// TIA Portal V21 export
// export: Created 2026-10-23T20:42:44.5110947Z, ExportSetting WithDefaults, DisplayName Totally Integrated Automation Portal, DisplayVersion V21 Update 1, DisplayName SINAMICS Startdrive Advanced, DisplayVersion V21 HF2, DisplayName SINAMICS Startdrive G110M, G120, G120C, G120D, G120P, G115D, DisplayVersion V21 HF2, DisplayName SINAMICS Startdrive G130, G150, S120, S150, G200, G220, S200, S210, S220, Innomotics MVD, DisplayVersion V21 HF2, DisplayName STEP 7 Professional, DisplayVersion V21 Update 1, DisplayName STEP 7 Safety, DisplayVersion V21, DisplayName Tech WebApplication, DisplayVersion V21, DisplayName WinCC Basic/Comfort/Advanced, DisplayVersion V21 Update 1, DisplayName WinCC Unified, DisplayVersion V21 Update 1
FUNCTION_BLOCK "FB_LadOpenBranch"   // FB8, LAD
TITLE = LAD open branch and parallel coils
{ S7_Optimized_Access := 'TRUE' }
VERSION : 0.1
// stored: AutoNumber true, IsIECCheckEnabled false, IsRetainMemResEnabled false, MemoryReserve 100, SetENOAutomatically false, UDAEnableTagReadback false
   VAR_INPUT
      Start : Bool;   // Start command
      Stop : Bool;   // Stop command
   END_VAR
   VAR_OUTPUT
      CoilA : Bool;   // First parallel coil
      CoilB : Bool;   // Second parallel coil
      CoilC : Bool;   // Third parallel coil, only without stop
      BranchOut : Bool;   // Coil of the network with the open branch
      StopLatched : Bool;   // Set by the open branch when stop is pressed during start
   END_VAR
   VAR
      StartCount : Int;   // Number of cycles with start pressed
   END_VAR
BEGIN

REGION Network 1: Several coils in parallel
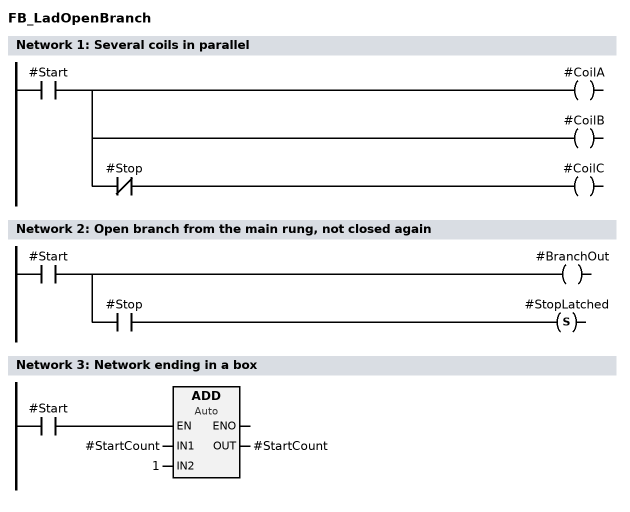
   RUNG wire#powerrail
      Contact( #Start )
      wire#w1
      Coil( #CoilA )
   END_RUNG
   RUNG wire#w1
      Coil( #CoilB )
   END_RUNG
   RUNG wire#w1
      I_Contact( #Stop )
      Coil( #CoilC )
   END_RUNG
   // the same network as SCL:
   #CoilA := #Start;
   #CoilB := #Start;
   #CoilC := #Start AND NOT #Stop;
END_REGION

REGION Network 2: Open branch from the main rung, not closed again
   RUNG wire#powerrail
      Contact( #Start )
      wire#w1
      Coil( #BranchOut )
   END_RUNG
   RUNG wire#w1
      Contact( #Stop )
      S_Coil( #StopLatched )
   END_RUNG
   // the same network as SCL:
   #BranchOut := #Start;
   IF #Start AND #Stop THEN #StopLatched := TRUE; END_IF;
END_REGION

REGION Network 3: Network ending in a box
   RUNG wire#powerrail
      Contact( #Start )
      Add(in1 := #StartCount, in2 := 1, out => #StartCount)
   END_RUNG
   // the same network as SCL:
   IF #Start THEN #StartCount := #StartCount + 1; END_IF;
END_REGION
END_FUNCTION_BLOCK
